PROGRAM Gr05MachineMode
VAR_INPUT
	(* Input variables / Eingang Variablen *)
	bEnable					:BOOL;						(* Enable Gr05MachineMode *)
END_VAR
VAR
	(* Enummerations *)

	(* Variables *)

	(* References *)

	(* Interfaces *)

	(* Instances *)

END_VAR

IF NOT bEnable
THEN
	RETURN;
END_IF;

Gr05Auto(bEnable := TRUE);			(* Call Program *)
Gr05Home(bEnable := TRUE);			(* Call Program *)
Gr05Manual(bEnable := TRUE);			(* Call Program *)

END_PROGRAM

(* stored: Version 1.1.0.1, ProductVersion 3.1.4024.15
   POU Gr05MachineMode: Id {f27b6dde-c85b-4fab-8a9a-7357614cef6d}, SpecialFunc None *)
